Staubli VAL3: insertPiston.pgx

program insertPiston()
// Level 3: four taught piston slots with tool presence sensing and bounded assembly.
begin
  // ============================================================
  // 40-43. BUSCAR UN PISTON: REVISAR SIEMPRE LOS 4 HUECOS DESDE EL 0
  // ============================================================
  // En cada montaje se recorre pistonIndex = 0,1,2,3 y se coge el
  // PRIMER hueco donde bIn0 detecta piston. partIndex solo cuenta montajes.
  // bIn0 esta en un LATERAL de la pinza y detecta presencia, no agarre.
  // Por hueco (todo con tTip):
  //   40 movej jCheckApproach (check + checkLift, calculado en start)
  //      movel jPistonCheck (ENSENADA) -> 41 leer bIn0
  //   Si NO hay piston: no se retira; se va directo al siguiente hueco.
  //   Si hay piston: 42 subir a jCheckApproach, ir al approach del pick,
  //      bajar vertical a jPistonPick, cerrar y subir al approach.
  // Si los 4 estan vacios: subir, avisar, esperar 2 s y repetir desde 0.
  pistonFound = false
  if physicalRun
    open(tTip)
  else
    delay(tTip.otime)
  endIf
  while !pistonFound
    pistonIndex = 0
    while !pistonFound and pistonIndex < 4
      cycleStep = 40
      putln("40 - Check piston slot (0..3):")
      putln(pistonIndex)
      putln("DBG 40A - movej to check approach")
      movej(jCheckApproach[pistonIndex], tTip, mNomSpeed)
      waitEndMove()
      putln("DBG 40B - movel to taught sensing pose jPistonCheck")
      movel(jointToPoint(tTip, world, jPistonCheck[pistonIndex]), tTip, mApproachSpeed)
      waitEndMove()
      cycleStep = 41
      pistonChecked = false
      if physicalRun
        // Asentar la herramienta y dejar actualizar physicalIO antes de leer.
        delay(0.15)
      else
        putln("MANUAL: set pistonPresent, then pistonChecked=true")
        wait(pistonChecked == true)
      endIf
      // Guardar la lectura ANTES de mover: physicalIO sigue refrescando
      // pistonPresent y al alejarse el sensor dejaria de verlo.
      pistonFound = pistonPresent
      putln("41 - Tool presence sensor bIn0:")
      if pistonFound
        putln("pistonPresent = true")
      else
        putln("pistonPresent = false")
        cycleStep = 43
        putln("43 - Empty slot; go to next slot")
        pistonIndex = pistonIndex + 1
      endIf
    endWhile
    if !pistonFound
      // Ultimo check fue el hueco 3: subir antes de volver al hueco 0.
      movel(jointToPoint(tTip, world, jCheckApproach[3]), tTip, mApproachSpeed)
      waitEndMove()
      putln("No piston in any slot; refill tray. Rescanning in 2 s.")
      delay(2)
    endIf
  endWhile

  // pistonIndex = primer hueco con piston detectado.
  cycleStep = 42
  putln("42 - Piston found; pick slot (0..3):")
  putln(pistonIndex)
  putln("DBG 42A - movel up to check approach")
  movel(jointToPoint(tTip, world, jCheckApproach[pistonIndex]), tTip, mApproachSpeed)
  waitEndMove()
  putln("DBG 42B - movel to pick approach")
  movel(jointToPoint(tTip, world, jPistonPick[2*pistonIndex]), tTip, mApproachSpeed)
  waitEndMove()
  putln("DBG 42C - movel down to pick; then close tTip")
  movel(jointToPoint(tTip, world, jPistonPick[2*pistonIndex+1]), tTip, mApproachSpeed)
  waitEndMove()
  if physicalRun
    close(tTip)
  else
    delay(tTip.ctime)
  endIf
  putln("DBG 42D - Piston gripped; withdraw to pick approach")
  movel(jointToPoint(tTip, world, jPistonPick[2*pistonIndex]), tTip, mApproachSpeed)
  waitEndMove()

  // ============================================================
  // 50. INSERTAR EL PISTON Y SOLTARLO ANTES DE RETIRARSE
  // ============================================================
  // TODO SIMULACION: confirmar el orden [0]/[1] de gridpiston.
  // TODO FISICO: ajustar alineacion y profundidad de jPistonInsert[1].
  // Este movimiento es por posicion; no mide fuerza ni confirma montaje.
  cycleStep = 50
  putln("50 - Insert piston into cylinder")
  putln("DBG 50A - BEFORE movej: insertion approach [0]")
  movej(jPistonInsert[0], tTip, mNomSpeed)
  waitEndMove()
  putln("DBG 50B - Insertion approach reached")
  movej(jointToPoint(tTip, world, jPistonInsert[1]), tTip, mInsertSpeed)
  waitEndMove()
  putln("DBG 50C - Insertion reached with tTip; opening gripper")
  if physicalRun
    open(tTip)
  else
    delay(tTip.otime)
  endIf
  putln("DBG 50D - BEFORE withdrawal with tTip to jPistonInsert[0]")
  movej(jointToPoint(tTip, world, jPistonInsert[0]), tTip, mInsertSpeed)
  waitEndMove()
  putln("DBG 50E - Tip withdrawal completed")

  // ============================================================
  // 55. POSTURA INTERMEDIA ANTES DE RECOGER EL CONJUNTO
  // ============================================================
  // Joint indicada por el usuario. Se alcanza DESPUES de soltar
  // el piston y retirarse con tTip, antes del agarre con tLateral.
  cycleStep = 55
  putln("DBG 55A - BEFORE movej: jAssemblyMove with tTip")
  movej(jAssemblyMove, tTip, mNomSpeed)
  waitEndMove()
  putln("DBG 55B - Assembly transit posture reached")

end
